FUNCTION_BLOCK AIS_TO_AIWS (* Composite FB for converting AIS (STRING) adapter to AIWS (WSTRING) adapter *)
  (* Standard: 61499-2; Description: Copyright (c) 2026 HR Agrartechnik GmbH This program and the accompanying materials are made available under the terms of the Eclipse Public License 2.0 which is available at https://www.eclipse.org/legal/epl-2.0/ SPDX-License-Identifier: EPL-2.0 *)
  (* Version 1.0, 2026-11-13, Franz Höpfinger, HR Agrartechnik GmbH, Initial Version - Luecke in der Adapter-Familie geschlossen *)
  PACKAGE adapter::conversion::unidirectional;
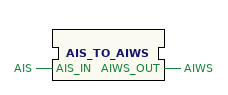
  SOCKETS
    AIS_IN : adapter::types::unidirectional::AIS; (* STRING Adapter Input *)
  END_SOCKETS
  PLUGS
    AIWS_OUT : adapter::types::unidirectional::AIWS; (* WSTRING Adapter Output *)
  END_PLUGS
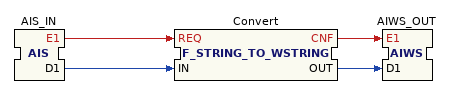
  FBS
    Convert : iec61131::conversion::F_STRING_TO_WSTRING;
  END_FBS
  EVENT_CONNECTIONS
    AIS_IN.E1 TO Convert.REQ;
    Convert.CNF TO AIWS_OUT.E1;
  END_CONNECTIONS
  DATA_CONNECTIONS
    AIS_IN.D1 TO Convert.IN;
    Convert.OUT TO AIWS_OUT.D1;
  END_CONNECTIONS
END_FUNCTION_BLOCK
